Staubli VAL3: seMaxJntForce.pgx

program seMaxJntForce()
  local num i
begin
//  if sArmType=="4_Axis"
//    for i=0 to 3
//      libTqe:tArm4Force[sArmDetail].nMaxJnt4Force[i]=nMaxJntForec[i]
//    endFor
//  elseIf sArmType=="6_Axis"
//    for i=0 to 5
//      libTqe:tArm6Force[sArmDetail].nMaxJnt6Force[i]=nMaxJntForec[i]
//    endFor
//  endIf
//  libTqe:libSave()
//  delay(0.1)
end
